// TIA Portal V21 export
// export: Created 2026-11-10T07:35:17.5081524Z, ExportSetting WithDefaults, DisplayName Totally Integrated Automation Portal, DisplayVersion V21 Update 3, DisplayName STEP 7 Professional, DisplayVersion V21 Update 3, DisplayName STEP 7 Safety, DisplayVersion V21, DisplayName Tech WebApplication, DisplayVersion V21, DisplayName WinCC Basic/Comfort/Advanced, DisplayVersion V21 Update 3, DisplayName WinCC Unified, DisplayVersion V21 Update 3
FUNCTION_BLOCK "FB_Lad_ex129"   // FB102, LAD
{ S7_Optimized_Access := 'TRUE' }
VERSION : 0.1
// stored: AutoNumber true, IsIECCheckEnabled false, IsRetainMemResEnabled false, MemoryReserve 100, SetENOAutomatically false, UDAEnableTagReadback false
   VAR_INPUT
      v_req : Bool;
      v_laddr : HW_DEVICE;
      v_detail : HW_SUBMODULE;
      v_mode : UInt;
   END_VAR
   VAR_OUTPUT
      v_done : Bool;
      v_busy : Bool;
      v_error : Bool;
      v_status : Word;
   END_VAR
   VAR_IN_OUT
      v_data : Array[0..99] of Byte;
   END_VAR
   VAR
      inst { S7_SetPoint := 'True'} : GetStationInfo;
   END_VAR
BEGIN

REGION Network 1: GetStationInfo - Read information of an IO device
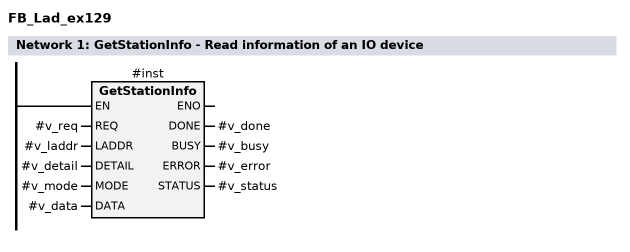
   RUNG wire#powerrail
      #inst.GetStationInfo(REQ := #v_req, LADDR := #v_laddr, DETAIL := #v_detail, MODE := #v_mode, DATA := #v_data, DONE => #v_done, BUSY => #v_busy, ERROR => #v_error, STATUS => #v_status)
   END_RUNG
   // the same network as SCL:
   #inst(REQ := #v_req,   // GetStationInfo
         LADDR := #v_laddr,
         DETAIL := #v_detail,
         MODE := #v_mode,
         DATA := #v_data,
         DONE => #v_done,
         BUSY => #v_busy,
         ERROR => #v_error,
         STATUS => #v_status);
END_REGION
END_FUNCTION_BLOCK
